SYSTEM System (* System Configuration *)
  (* Standard: 61499-1 *)
  (* Version 0.0, 9/9/2026, lizar, Schneider Electric *)
  {SET_ATTRIBUTE(System.Device.FolderPath, EcoRT_0)}
  APPLICATION APP1
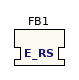
    FBS
      FB1 : E_RS;
    END_FBS
  END_APPLICATION
  APPLICATION E_TRAIN_TEST
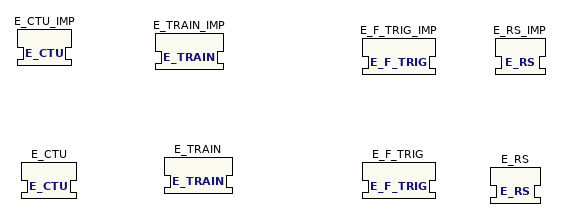
    FBS
      E_TRAIN_IMP : E_TRAIN;
      E_TRAIN : E_TRAIN;
      E_F_TRIG_IMP : E_F_TRIG;
      E_F_TRIG : E_F_TRIG;
      E_CTU_IMP : E_CTU;
      E_CTU : E_CTU;
      E_RS : E_RS;
      E_RS_IMP : E_RS;
    END_FBS
  END_APPLICATION
  DEVICE EcoRT_0 : Soft_dPAC
    RESOURCE RES0 : EMB_RES_ECO
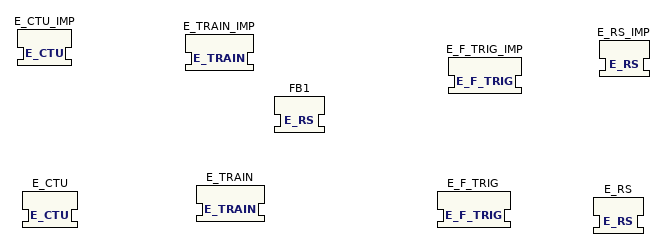
      FBS
        FB1 : E_RS;
        E_TRAIN_IMP : E_TRAIN;
        E_TRAIN : E_TRAIN;
        E_F_TRIG_IMP : E_F_TRIG;
        E_F_TRIG : E_F_TRIG;
        E_CTU_IMP : E_CTU;
        E_CTU : E_CTU;
        E_RS_IMP : E_RS;
        E_RS : E_RS;
      END_FBS
    END_RESOURCE
  END_DEVICE
  MAPPINGS
    APP1.FB1 ON EcoRT_0.RES0;
    E_TRAIN_TEST.E_TRAIN_IMP ON EcoRT_0.RES0;
    E_TRAIN_TEST.E_TRAIN ON EcoRT_0.RES0;
    E_TRAIN_TEST.E_F_TRIG_IMP ON EcoRT_0.RES0;
    E_TRAIN_TEST.E_F_TRIG ON EcoRT_0.RES0;
    E_TRAIN_TEST.E_CTU_IMP ON EcoRT_0.RES0;
    E_TRAIN_TEST.E_CTU ON EcoRT_0.RES0;
    E_TRAIN_TEST.E_RS_IMP ON EcoRT_0.RES0;
    E_TRAIN_TEST.E_RS ON EcoRT_0.RES0;
  END_MAPPINGS
END_SYSTEM
(* other elements stored in the file *)
(* Layer Name=RS_Test *)
(* FBName Name=FB1 *)
